(* IEC 61131-3 sources: st2fb/corpus_hard/unsupported_st/u03_tank_strapping, 2 files *)

(* ---- control_flat.st ---- *)
(* Solvability control, never shown to a model: the same behaviour in the translator's v1 subset. The table became
   a chain of IFs, and RETURN became an enclosing IF. *)
FUNCTION_BLOCK TANK_STRAPPING
VAR_INPUT
  LEVEL_MM : REAL;
  DENSITY : REAL;
  HOLD : BOOL;
END_VAR
VAR_OUTPUT
  VOLUME_L : REAL;
  MASS_KG : DINT;
  SEGMENT : INT;
  OUT_OF_RANGE : BOOL;
END_VAR
VAR
  L0, L1, V0, V1 : REAL;
  FRACTION : REAL;
END_VAR
  IF NOT HOLD THEN
    OUT_OF_RANGE := (LEVEL_MM < 0.0) OR (LEVEL_MM > 2000.0);
    IF LEVEL_MM <= 200.0 THEN
      SEGMENT := 0;
      L0 := 0.0;
      L1 := 200.0;
      V0 := 0.0;
      V1 := 150.0;
    ELSIF LEVEL_MM <= 400.0 THEN
      SEGMENT := 1;
      L0 := 200.0;
      L1 := 400.0;
      V0 := 150.0;
      V1 := 340.0;
    ELSIF LEVEL_MM <= 800.0 THEN
      SEGMENT := 2;
      L0 := 400.0;
      L1 := 800.0;
      V0 := 340.0;
      V1 := 800.0;
    ELSIF LEVEL_MM <= 1200.0 THEN
      SEGMENT := 3;
      L0 := 800.0;
      L1 := 1200.0;
      V0 := 800.0;
      V1 := 1350.0;
    ELSE
      SEGMENT := 4;
      L0 := 1200.0;
      L1 := 2000.0;
      V0 := 1350.0;
      V1 := 2600.0;
    END_IF;
    FRACTION := (LEVEL_MM - L0) / (L1 - L0);
    FRACTION := LIMIT(0.0, FRACTION, 1.0);
    VOLUME_L := V0 + FRACTION * (V1 - V0);
    MASS_KG := REAL_TO_DINT(VOLUME_L * DENSITY);
  END_IF;
END_FUNCTION_BLOCK

(* ---- program.st ---- *)
(* Tank strapping table: level to volume by linear interpolation. *)
TYPE
  STRAP_TABLE : ARRAY[0..5] OF REAL;
END_TYPE

FUNCTION_BLOCK TANK_STRAPPING
VAR_INPUT
  LEVEL_MM : REAL;
  DENSITY : REAL;
  HOLD : BOOL;
END_VAR
VAR_OUTPUT
  VOLUME_L : REAL;
  MASS_KG : DINT;
  SEGMENT : INT;
  OUT_OF_RANGE : BOOL;
END_VAR
VAR
  LEVELS : STRAP_TABLE := [0.0, 200.0, 400.0, 800.0, 1200.0, 2000.0];
  VOLUMES : STRAP_TABLE := [0.0, 150.0, 340.0, 800.0, 1350.0, 2600.0];
  I : INT;
  FRACTION : REAL;
END_VAR
  IF HOLD THEN
    RETURN;
  END_IF;
  OUT_OF_RANGE := (LEVEL_MM < LEVELS[0]) OR (LEVEL_MM > LEVELS[5]);
  I := 0;
  REPEAT
    IF LEVEL_MM <= LEVELS[I + 1] THEN
      EXIT;
    END_IF;
    I := I + 1;
  UNTIL I >= 4
  END_REPEAT;
  SEGMENT := I;
  FRACTION := (LEVEL_MM - LEVELS[I]) / (LEVELS[I + 1] - LEVELS[I]);
  FRACTION := LIMIT(0.0, FRACTION, 1.0);
  VOLUME_L := VOLUMES[I] + FRACTION * (VOLUMES[I + 1] - VOLUMES[I]);
  MASS_KG := REAL_TO_DINT(VOLUME_L * DENSITY);
END_FUNCTION_BLOCK
